Fanuc KAREL source: ka00155.KL

-- PROVISIONAL review KL for V940-1; original PC SHA256 f2e81668cfa7df35c2a13bf2fcc13463b14c6a1d801d3c4fa09a3434a7b8cd30
-- Incomplete behavior may be omitted. Consult companion uncertainty JSON. Do not deploy.
PROGRAM KA00155
%NOLOCKGROUP
-- UNRESOLVED_DECL SRC type=002011
-- UNRESOLVED_DECL DST type=002011
BEGIN
  -- V9_COMPOSED_GLOBAL_TRANSFER_HINT repetitions=1; address IDs observed; pairing/direction/source/runtime held
  -- V9_TWO_GLOBAL_ADDRESS_COPY_HINT bounded five-record physical form; type/direction/source/runtime held
  -- V9_ZERO_TABLE_METADATA_HINT layout=0001; no indexed target words; source/name/runtime held
  -- UNRESOLVED_PC offsets 5-19; opcodes 22,22,1E
  -- UNRESOLVED_PC offsets 24-28; opcodes 7F
END KA00155
